Fanuc KAREL source: ko00044.KL

-- PROVISIONAL review KL for V1013-1; original PC SHA256 d9276e01b97fdc7eb811bc9a5bf02202f136e87517f9d16853d55d39a39ad56c
-- Incomplete behavior may be omitted. Consult companion uncertainty JSON. Do not deploy.
PROGRAM KO00044
%NOLOCKGROUP
BEGIN
  -- UNRESOLVED_PC offsets 5-12; opcodes 9D,23
  -- UNRESOLVED_PC offsets 17-69; opcodes 27,27,49,7E,AD,27,49,7E,AD,22,31,7E,4A
  -- UNRESOLVED_PC offsets 74-78; opcodes 7F
END KO00044
